(* IEC 61131-3 sources: plc-iiot-stack/tests/POUs/FB_MqttTelemetry_Test, 13 files *)

(* ---- BudgetLimitsPublishesPerCallRoundRobin.method.decl.st ---- *)
// Не больше uiMaxPerCycle за вызов, остальные — в следующих, по кругу.
METHOD PRIVATE BudgetLimitsPublishesPerCallRoundRobin
VAR_INST
    fbFake : FB_MqttClientFake;
    fbTel : FB_MqttTelemetry;
    aPts : ARRAY[1..5] OF ST_IiotPoint;
END_VAR

(* ---- ClientRefusalIsCountedAndRetried.method.decl.st ---- *)
// Клиент не принял — udiFailed, метрики ждут и уходят позже.
METHOD PRIVATE ClientRefusalIsCountedAndRetried
VAR_INST
    fbFake : FB_MqttClientFake;
    fbTel : FB_MqttTelemetry;
    aPts : ARRAY[1..4] OF ST_IiotPoint;
END_VAR

(* ---- DeadbandAndMinInterval.method.decl.st ---- *)
// Зона нечувствительности и не чаще раза в секунду на метрику.
METHOD PRIVATE DeadbandAndMinInterval
VAR_INST
    fbFake : FB_MqttClientFake;
    fbTel : FB_MqttTelemetry;
    aPts : ARRAY[1..4] OF ST_IiotPoint;
END_VAR

(* ---- IntegerAnyChangeAndPeriodicOnly.method.decl.st ---- *)
// Целые — при любом изменении; время работы узла — только контрольно.
METHOD PRIVATE IntegerAnyChangeAndPeriodicOnly
VAR_INST
    fbFake : FB_MqttClientFake;
    fbTel : FB_MqttTelemetry;
    aPts : ARRAY[1..4] OF ST_IiotPoint;
END_VAR

(* ---- NegativeAndLargeValues.method.decl.st ---- *)
// Отрицательное Analog и большой счётчик Integer — без потери знака и разрядов.
METHOD PRIVATE NegativeAndLargeValues
VAR_INST
    fbFake : FB_MqttClientFake;
    fbTel : FB_MqttTelemetry;
    aPts : ARRAY[1..4] OF ST_IiotPoint;
END_VAR

(* ---- NotFiniteValueSendsLastFiniteAsBad.method.decl.st ---- *)
// Значение стало NaN: схема требует число — передаётся последнее опубликованное конечное значение с
// quality = bad; конечное значение возвращает исходное качество.
METHOD PRIVATE NotFiniteValueSendsLastFiniteAsBad
VAR_INST
    fbFake : FB_MqttClientFake;
    fbTel : FB_MqttTelemetry;
    aPts : ARRAY[1..4] OF ST_IiotPoint;
END_VAR
VAR
    lwNan : LWORD := 16#7FF8000000000000;
    pBits : POINTER TO LREAL;
END_VAR

(* ---- PeriodRepublishesAll.method.decl.st ---- *)
// По истечении периода — все метрики, раньше — нет.
METHOD PRIVATE PeriodRepublishesAll
VAR_INST
    fbFake : FB_MqttClientFake;
    fbTel : FB_MqttTelemetry;
    aPts : ARRAY[1..4] OF ST_IiotPoint;
END_VAR

(* ---- PublishesAllAfterBirthWithExactJson.method.decl.st ---- *)
// После рождения узла — все метрики; точный JSON, QoS 1, retain.
METHOD PRIVATE PublishesAllAfterBirthWithExactJson
VAR_INST
    fbFake : FB_MqttClientFake;
    fbTel : FB_MqttTelemetry;
    aPts : ARRAY[1..4] OF ST_IiotPoint;
END_VAR

(* ---- QualityChangeIsImmediate.method.decl.st ---- *)
// Смена качества публикуется сразу, без ожидания интервала.
METHOD PRIVATE QualityChangeIsImmediate
VAR_INST
    fbFake : FB_MqttClientFake;
    fbTel : FB_MqttTelemetry;
    aPts : ARRAY[1..4] OF ST_IiotPoint;
END_VAR

(* ---- RepublishesAllAfterReconnect.method.decl.st ---- *)
// Связь пропала и вернулась с новым рождением — все метрики заново.
METHOD PRIVATE RepublishesAllAfterReconnect
VAR_INST
    fbFake : FB_MqttClientFake;
    fbTel : FB_MqttTelemetry;
    aPts : ARRAY[1..4] OF ST_IiotPoint;
END_VAR

(* ---- Run.method.decl.st ---- *)
// Вызов FB_MqttTelemetry: префикс vodokanal/kns1/station, ts 1792137600250, период 10 с.
METHOD PRIVATE Run
VAR_IN_OUT
    fbTelemetry : FB_MqttTelemetry;
    fbClient : FB_MqttClientFake;
    aPointTable : ARRAY[*] OF ST_IiotPoint;
END_VAR
VAR_INPUT
    ltAt : LTIME;
    xReadyIn : BOOL;
END_VAR

(* ---- Setup.method.decl.st ---- *)
// Четыре метрики: уровень (Analog, зона 0.01 м), работа насоса (Integer), пуски (Integer), время работы узла
// (только контрольно); связь есть.
METHOD PRIVATE Setup
VAR_IN_OUT
    fbClient : FB_MqttClientFake;
    aPointTable : ARRAY[1..4] OF ST_IiotPoint;
END_VAR

(* ---- WaitsForBirthAndClock.method.decl.st ---- *)
// До рождения узла и без часов ПЛК — ничего; потом — всё.
METHOD PRIVATE WaitsForBirthAndClock
VAR_INST
    fbFake : FB_MqttClientFake;
    fbTel : FB_MqttTelemetry;
    aPts : ARRAY[1..4] OF ST_IiotPoint;
END_VAR
